// TIA Portal V21 export
// export: Created 2026-10-23T20:43:24.2078009Z, ExportSetting WithDefaults, DisplayName Totally Integrated Automation Portal, DisplayVersion V21 Update 1, DisplayName SINAMICS Startdrive Advanced, DisplayVersion V21 HF2, DisplayName SINAMICS Startdrive G110M, G120, G120C, G120D, G120P, G115D, DisplayVersion V21 HF2, DisplayName SINAMICS Startdrive G130, G150, S120, S150, G200, G220, S200, S210, S220, Innomotics MVD, DisplayVersion V21 HF2, DisplayName STEP 7 Professional, DisplayVersion V21 Update 1, DisplayName STEP 7 Safety, DisplayVersion V21, DisplayName Tech WebApplication, DisplayVersion V21, DisplayName WinCC Basic/Comfort/Advanced, DisplayVersion V21 Update 1, DisplayName WinCC Unified, DisplayVersion V21 Update 1
FUNCTION_BLOCK "FB_AnaUnused"   // FB15, SCL
TITLE = Analyzer: unused variables
{ S7_Optimized_Access := 'TRUE' }
VERSION : 0.1
// Rule C26j: UnusedInput, UnusedStatic and UnusedTemp are never used
// stored: AutoNumber true, IsIECCheckEnabled false, IsRetainMemResEnabled false, MemoryReserve 100, SetENOAutomatically false, UDAEnableTagReadback false
   VAR_INPUT
      UsedInput : Int;   // Used input
      UnusedInput : Int;   // Unused input
   END_VAR
   VAR_OUTPUT
      Result : Int;   // Result
   END_VAR
   VAR
      UnusedStatic : Int;   // Unused static variable
   END_VAR
   VAR_TEMP
      UnusedTemp : Int;   // Unused temporary variable
   END_VAR
BEGIN

       #Result := #UsedInput * 2;
END_FUNCTION_BLOCK
